FUNCTION_BLOCK FB_LimitAlarm
(*
	One high or low threshold alarm with deadband, on-delay and optional latching.
	High alarm: on when value >= threshold for delay, off when value < threshold - deadband.
	Low alarm:  on when value <= threshold for delay, off when value > threshold + deadband.
	A latched alarm stays on until reset is TRUE and the condition has cleared.
*)
VAR_INPUT
	value				: LREAL; //value to check
	threshold				: LREAL; //alarm threshold
	highAlarm			: BOOL; //TRUE = high alarm, FALSE = low alarm
	enable				: BOOL; //alarm is enabled
	deadband			: LREAL; //hysteresis before the condition clears
	delay				: TIME; //condition must be present this long before the alarm turns on
	latch				: BOOL; //alarm stays on until reset
	reset				: BOOL; //reset a latched alarm (only clears once the condition is gone)
END_VAR
VAR_OUTPUT
	active				: BOOL; //alarm is on
	condition			: BOOL; //threshold currently exceeded (before delay and latch)
END_VAR
VAR
	//Timers
	delayTimer			: TON; //on-delay
END_VAR

Evaluate();

METHOD PROTECTED Evaluate
//Condition with hysteresis
IF highAlarm THEN
	IF value >= threshold THEN
		condition := TRUE;
	ELSIF value < threshold - deadband THEN
		condition := FALSE;
	END_IF
ELSE
	IF value <= threshold THEN
		condition := TRUE;
	ELSIF value > threshold + deadband THEN
		condition := FALSE;
	END_IF
END_IF
condition := condition AND enable;

delayTimer(IN := condition, PT := delay);

IF latch THEN
	active S= delayTimer.Q;
	active R= reset AND NOT condition;
ELSE
	active := delayTimer.Q;
END_IF
END_METHOD

END_FUNCTION_BLOCK

(* stored: Version 1.1.0.1, ProductVersion 3.1.4024.12
   POU FB_LimitAlarm: Id {15488189-7294-462f-928a-2f67960bcc3c}, SpecialFunc None
   Folder Protected: Id {64e04b85-2af5-4e59-bd1f-4b66773f093e}
   Folder Logic: Id {83f228a0-9d67-4dd5-a5b7-4109f83af035}
   Method Evaluate: Id {40fc6caa-278e-4531-b941-eb67b60b5ac4} *)
